// TIA Portal V20 export
DATA_BLOCK "03_Betriebsart_DB"   // DB11
// stored: InstanceOfName 03_Betriebsart, InstanceOfType FB
"03_Betriebsart"
   // VAR
   //    Projektnummer : WString;
   //    Projektname : WString;
   //    Validierung_Datum : WString;
   //    Validierung_Name : WString;
   //    Validierung_F_PROG_SIG : DWord;
   //    Aktuell_F_PROG_SIG : DWord;
   //    F_PROG_SIG_stimmt_überein : Bool;
   //    Simulation_aktiv : Bool;
   //    IN_Betriebsart_Manuell { ExternalAccessible := 'False'; ExternalVisible := 'False'; ExternalWritable := 'False'} : Bool;
   //    BA_Automatik_HMFP : Bool;
   //    BA_Automatik_FP : Bool;
   //    IN_Betriebsart_Automatik { ExternalAccessible := 'False'; ExternalVisible := 'False'; ExternalWritable := 'False'} : Bool;
   //    BA_Verwaltung_HMFP : Bool;
   //    BA_Verwaltung_FP : Bool;
   //    IN_Betriebsart_Verwaltung { ExternalAccessible := 'False'; ExternalVisible := 'False'; ExternalWritable := 'False'} : Bool;
   //    IN_Betriebsart_Richten { ExternalAccessible := 'False'; ExternalVisible := 'False'; ExternalWritable := 'False'} : Bool;
   //    Systemdruck_OK : Bool;
   //    Betriebsart : Int;
   //    BA_Manuell_HMFP : Bool;
   //    BA_Manuell_FP : Bool;
   //    BA_Manuell : Bool;
   //    BA_Automatik : Bool;
   //    BA_Verwaltung : Bool;
   //    BA_Richten_HMFP : Bool;
   //    BA_Richten_FP : Bool;
   //    BA_Richten : Bool;
   //    BA_0 : Bool;
   //    BA_0_HMFP : Bool;
   //    BA_0_FP : Bool;
   //    BA_0_groesser_1_5 : Bool;
   //    TON_BA_0_groesser_1_5 { S7_SetPoint := 'True'} : TON_TIME;
   //    TON_Rücksetzen_der_Betriebsart { S7_SetPoint := 'True'} : TON_TIME;
   //    TON_Türen_setzen_zum_öffnen { S7_SetPoint := 'True'} : TON_TIME;
   //    "TOF_MRW Not-Halt Überwachung deaktivieren" { S7_SetPoint := 'True'} : TOF_TIME;
   //    HM_MRW_Zeitverzögerung { S7_SetPoint := 'True'} : Bool;
   //    Türen_sind_verriegelt { S7_SetPoint := 'True'} : Bool;
   //    "NOT-HALT OK" : Bool;
   //    "NOT-HALT_HMFN" : Bool;
   //    "NOT-HALT_FN" : Bool;
   //    Start_Taste : Bool;
   //    Start_Taste_HMFP : Bool;
   //    Start_Taste_FP : Bool;
   //    ACK_Taste : Bool;
   //    ACK_Taste_HMFP : Bool;
   //    ACK_Taste_FP : Bool;
   //    Stopp_Taste : Bool;
   //    "Schutztüren OK" : Bool;
   //    Schutztüren_HMFN : Bool;
   //    Schutztüren_FN : Bool;
   //    Schutztüren_HMFP : Bool;
   //    Schutztüren_FP : Bool;
   //    "Druckbereich entlüftet" : Bool;
   //    Antriebe_sicher : Bool;
   //    Zuhaltung_Freigeben : Bool;
   //    Roboter_Motor_Ein : Bool;
   //    "P_Trig_Betriebsart Manuell" : Bool;
   //    "P_Trig_Betriebsart Automatik" : Bool;
   //    "P_Trig_Betriebsart Verwaltung" : Bool;
   //    "P_Trig_Betriebsart Richten" : Bool;
   //    TON_Hauptventil_aus { S7_SetPoint := 'True'} : TON_TIME;
   //    TON_Hauptventil_aus_status_Reset { S7_SetPoint := 'True'} : TON_TIME;
   //    Flanke_Hauptventil_aus { S7_SetPoint := 'True'} : Bool;
   //    Hauptventil_Reset : Bool;
   //    KP8_Bedienerkonsole { S7_SetPoint := 'True'} : "KP8";
   // END_VAR
BEGIN
END_DATA_BLOCK
